// TIA Portal V20 export
Screen "190RB06_J5"  1276x673
  ScreenItem "Graphic view_2" at 277,106 size 704x526  Type=HmiGraphicView
  ScreenItem "Line_Header_X0_Y64" at -3,67 size 1276x0  Type=HmiLine
  ScreenItem "permanentareaborderrectangle" at 0,0 size 0x0  Type=HmiRectangle
  ScreenItem "Button_Back" at 2,2 size 90x60  Type=HmiButton
  ScreenItem "Fusszeile_Button_ManualOPMode1_4" at 1181,2 size 90x60  Type=HmiButton
  ScreenItem "Title_ScreenOverview_X390_Y2_5" at 393,4 size 510x57  Type=HmiTextBox
  ScreenItem "Fusszeile_Button_ManualOPMode1_1" at 1088,2 size 90x60  Type=HmiButton
  ScreenItem "Title_ScreenOverview_X390_Y2_1" at 1138,86 size 139x57  Type=HmiTextBox
  ScreenItem "Title_ScreenOverview_X390_Y2_6" at 1138,152 size 139x57  Type=HmiTextBox
  ScreenItem "Title_ScreenOverview_X390_Y2_7" at 1138,152 size 139x57  Type=HmiTextBox
  ScreenItem "文本域_15" at 397,174 size 140x20  Type=HmiTextBox
  ScreenItem "Line_16" at 458,254 size 24x110  Type=HmiLine
  ScreenItem "Line_4" at 956,205 size 41x13  Type=HmiLine
  ScreenItem "文本域_11" at 1001,173 size 134x40  Type=HmiTextBox
  ScreenItem "Line_2" at 863,272 size 130x24  Type=HmiLine
  ScreenItem "Line_3" at 847,338 size 142x12  Type=HmiLine
  ScreenItem "文本域_4" at 985,415 size 134x40  Type=HmiTextBox
  ScreenItem "Line_5" at 870,375 size 115x56  Type=HmiLine
  ScreenItem "文本域_5" at 985,548 size 134x40  Type=HmiTextBox
  ScreenItem "Line_6" at 794,574 size 177x14  Type=HmiLine
  ScreenItem "文本域_6" at 624,574 size 134x40  Type=HmiTextBox
  ScreenItem "Line_7" at 606,577 size 13x20  Type=HmiLine
  ScreenItem "Line_8" at 512,488 size 14x45  Type=HmiLine
  ScreenItem "文本域_7" at 440,537 size 134x40  Type=HmiTextBox
  ScreenItem "Line_9" at 267,592 size 77x8  Type=HmiLine
  ScreenItem "文本域_8" at 128,568 size 134x40  Type=HmiTextBox
  ScreenItem "文本域_9" at 20,516 size 134x40  Type=HmiTextBox
  ScreenItem "Line_10" at 159,485 size 140x63  Type=HmiLine
  ScreenItem "Line_11" at 180,436 size 156x16  Type=HmiLine
  ScreenItem "文本域_12" at 30,335 size 134x40  Type=HmiTextBox
  ScreenItem "Line_12" at 172,365 size 186x2  Type=HmiLine
  ScreenItem "Line_13" at 184,262 size 201x77  Type=HmiLine
  ScreenItem "文本域_14" at 472,77 size 134x40  Type=HmiTextBox
  ScreenItem "Line_14" at 534,164 size 16x101  Type=HmiLine
  ScreenItem "文本域_16" at 77,90 size 134x40  Type=HmiTextBox
  ScreenItem "Line_15" at 219,134 size 127x27  Type=HmiLine
  ScreenItem "文本域_17" at 643,480 size 140x20  Type=HmiTextBox
  ScreenItem "Line_17" at 715,363 size 0x111  Type=HmiLine
  ScreenItem "文本域_1" at 646,200 size 120x20  Type=HmiTextBox
  ScreenItem "Line_1" at 611,220 size 30x24  Type=HmiLine
  ScreenItem "文本域_18" at 635,77 size 134x40  Type=HmiTextBox
  ScreenItem "Line_18" at 612,130 size 35x38  Type=HmiLine
  ScreenItem "文本域_19" at 850,95 size 134x40  Type=HmiTextBox
  ScreenItem "Line_19" at 797,143 size 68x20  Type=HmiLine
  ScreenItem "Title_ScreenOverview_X390_Y2_44" at 121,134 size 52x19  Type=HmiTextBox
  ScreenItem "Title_ScreenOverview_X390_Y2_45" at 121,154 size 25x21  Type=HmiTextBox
  ScreenItem "Title_ScreenOverview_X390_Y2_46" at 148,154 size 25x21  Type=HmiTextBox
  ScreenItem "Title_ScreenOverview_X390_Y2_2" at 513,117 size 52x19  Type=HmiTextBox
  ScreenItem "Title_ScreenOverview_X390_Y2_3" at 513,137 size 25x21  Type=HmiTextBox
  ScreenItem "Title_ScreenOverview_X390_Y2_4" at 540,137 size 25x21  Type=HmiTextBox
  ScreenItem "Title_ScreenOverview_X390_Y2_8" at 679,116 size 52x19  Type=HmiTextBox
  ScreenItem "Title_ScreenOverview_X390_Y2_9" at 679,136 size 25x21  Type=HmiTextBox
  ScreenItem "Title_ScreenOverview_X390_Y2_10" at 706,136 size 25x21  Type=HmiTextBox
  ScreenItem "Title_ScreenOverview_X390_Y2_11" at 891,135 size 52x19  Type=HmiTextBox
  ScreenItem "Title_ScreenOverview_X390_Y2_12" at 891,155 size 25x21  Type=HmiTextBox
  ScreenItem "Title_ScreenOverview_X390_Y2_13" at 918,155 size 25x21  Type=HmiTextBox
  ScreenItem "Title_ScreenOverview_X390_Y2_14" at 1044,213 size 52x19  Type=HmiTextBox
  ScreenItem "Title_ScreenOverview_X390_Y2_15" at 1044,233 size 25x21  Type=HmiTextBox
  ScreenItem "Title_ScreenOverview_X390_Y2_16" at 1071,233 size 25x21  Type=HmiTextBox
  ScreenItem "Title_ScreenOverview_X390_Y2_17" at 1024,455 size 52x19  Type=HmiTextBox
  ScreenItem "Title_ScreenOverview_X390_Y2_18" at 1024,475 size 25x21  Type=HmiTextBox
  ScreenItem "Title_ScreenOverview_X390_Y2_19" at 1051,475 size 25x21  Type=HmiTextBox
  ScreenItem "Title_ScreenOverview_X390_Y2_20" at 1024,592 size 52x19  Type=HmiTextBox
  ScreenItem "Title_ScreenOverview_X390_Y2_21" at 1024,612 size 25x21  Type=HmiTextBox
  ScreenItem "Title_ScreenOverview_X390_Y2_22" at 1051,612 size 25x21  Type=HmiTextBox
  ScreenItem "Title_ScreenOverview_X390_Y2_23" at 658,614 size 52x19  Type=HmiTextBox
  ScreenItem "Title_ScreenOverview_X390_Y2_24" at 658,634 size 25x21  Type=HmiTextBox
  ScreenItem "Title_ScreenOverview_X390_Y2_25" at 685,634 size 25x21  Type=HmiTextBox
  ScreenItem "Title_ScreenOverview_X390_Y2_26" at 482,581 size 52x19  Type=HmiTextBox
  ScreenItem "Title_ScreenOverview_X390_Y2_27" at 482,601 size 25x21  Type=HmiTextBox
  ScreenItem "Title_ScreenOverview_X390_Y2_28" at 509,601 size 25x21  Type=HmiTextBox
  ScreenItem "Title_ScreenOverview_X390_Y2_29" at 167,608 size 52x19  Type=HmiTextBox
  ScreenItem "Title_ScreenOverview_X390_Y2_30" at 167,628 size 25x21  Type=HmiTextBox
  ScreenItem "Title_ScreenOverview_X390_Y2_31" at 194,628 size 25x21  Type=HmiTextBox
  ScreenItem "Title_ScreenOverview_X390_Y2_32" at 50,561 size 52x19  Type=HmiTextBox
  ScreenItem "Title_ScreenOverview_X390_Y2_33" at 50,581 size 25x21  Type=HmiTextBox
  ScreenItem "Title_ScreenOverview_X390_Y2_34" at 77,581 size 25x21  Type=HmiTextBox
  ScreenItem "Title_ScreenOverview_X390_Y2_35" at 69,375 size 52x19  Type=HmiTextBox
  ScreenItem "Title_ScreenOverview_X390_Y2_36" at 69,395 size 25x21  Type=HmiTextBox
  ScreenItem "Title_ScreenOverview_X390_Y2_37" at 96,395 size 25x21  Type=HmiTextBox
  ScreenItem "Rectangle_13" at 0,0 size 165x48  Type=HmiRectangle
  ScreenItem "文本域_20" at 2,1 size 132x45  Type=HmiTextBox
  ScreenItem "圆_5" at 0,0 size 100x30  Type=HmiCircle
  ScreenItem "圆_6" at 0,0 size 100x30  Type=HmiCircle
  ScreenItem "Rectangle_1" at 0,0 size 141x48  Type=HmiRectangle
  ScreenItem "文本域_13" at 2,1 size 113x45  Type=HmiTextBox
  ScreenItem "圆_1" at 0,0 size 100x30  Type=HmiCircle
  ScreenItem "圆_2" at 0,0 size 100x30  Type=HmiCircle
  ScreenItem "Rectangle_2" at 0,0 size 141x48  Type=HmiRectangle
  ScreenItem "文本域_10" at 2,1 size 113x45  Type=HmiTextBox
  ScreenItem "圆_3" at 0,0 size 100x30  Type=HmiCircle
  ScreenItem "圆_4" at 0,0 size 100x30  Type=HmiCircle
  ScreenItem "Rectangle_3" at 0,0 size 165x48  Type=HmiRectangle
  ScreenItem "文本域_2" at 2,1 size 132x45  Type=HmiTextBox
  ScreenItem "圆_7" at 0,0 size 100x30  Type=HmiCircle
  ScreenItem "圆_8" at 0,0 size 100x30  Type=HmiCircle
